Fanuc KAREL source: KT00833.KL

PROGRAM KT00833
%NOLOCKGROUP
VAR
  I1: INTEGER
  I2: INTEGER
  OUT: REAL
BEGIN
  I1 = 2
  I2 = 3
  I1 = 2
  I2 = 3
  OUT = SQRT(I1)
END KT00833
